(* IEC 61131-3 sources: FACTORY_io/misiones/01-marcha-paro/proyecto/plc, 1 file *)

(* ---- program.st ---- *)
(* Misión 1 · Marcha y paro

   Objetivo: que el pulsador Marcha ponga en marcha la cinta y el alimentador de cajas, que sigan
   funcionando al soltarlo, y que Paro los detenga. Si se pulsan los dos a la vez, gana Paro.

   Las señales ya están declaradas con los nombres que usan las piezas de la escena.
   Escribe tu lógica debajo de la línea "Tu programa". *)

(* Cómo probarlo: pulsa Play (▶). Para accionar un pulsador, selecciónalo en la lista Scene
   (por ejemplo «Pulsador Marcha») y pulsa la tecla C. En la pestaña Watch ves las variables.
   Cuando creas que está, pulsa «Run tests» (junto a Play): es el juez de la misión. *)
VAR_INPUT
  FotocelulaSalida : BOOL;  (* fotocélula al final de la cinta: TRUE con caja delante *)
  Marcha : BOOL;            (* pulsador verde: TRUE solo mientras se pulsa *)
  Paro : BOOL;              (* pulsador rojo: TRUE solo mientras se pulsa *)
  CajasSalida : INT;        (* cajas retiradas por el sumidero *)
END_VAR
VAR_OUTPUT
  CintaMarcha : BOOL;       (* TRUE: la cinta se mueve *)
  Alimentador : BOOL;       (* TRUE: el alimentador suelta cajas *)
END_VAR
VAR
  (* tus variables internas *)
END_VAR

(* ---- Tu programa ---- *)
